(* IEC 61131-3 sources: model-first-plc-agent-ai/results/T2-W-09, 2 files *)

(* ---- a1_code.st ---- *)
FUNCTION_BLOCK TankFillingRuntime
VAR_INPUT
    start : BOOL;
    stop : BOOL;
    LSH : BOOL;
    LSHH : BOOL;
    TimerDuration : TIME;
END_VAR
VAR_OUTPUT
    fill_valve : BOOL;
    discharge_valve : BOOL;
END_VAR
VAR
    x0 : BOOL := TRUE;
    x1 : BOOL := FALSE;
    t1 : BOOL;
    t2 : BOOL;
    timer_done : BOOL := FALSE;
    FillingTimer : TON;
END_VAR

(* Evaluate the start transition from the current situation. *)
t1 := x0 AND start AND NOT stop AND NOT LSHH;

(* Start timing in the same scan that the filling step is entered. *)
FillingTimer(
    IN := x1 OR t1,
    PT := TimerDuration
);

(* The owned condition is neutral on entry to x1. *)
timer_done := x1 AND FillingTimer.Q;

(* Evaluate the return transition before updating the situation. *)
t2 := x1 AND (stop OR LSHH OR timer_done);

IF t1 THEN
    x0 := FALSE;
    x1 := TRUE;
ELSIF t2 THEN
    x0 := TRUE;
    x1 := FALSE;
END_IF;

(* Reset the owned timer immediately when its step is inactive. *)
IF NOT x1 THEN
    FillingTimer(IN := FALSE, PT := TimerDuration);
    timer_done := FALSE;
END_IF;

fill_valve := x1;
discharge_valve := FALSE;

END_FUNCTION_BLOCK

PROGRAM Main
VAR
    StartCommand AT %IX100.0 : BOOL;
    StopCommand AT %IX100.1 : BOOL;
    LSH AT %IX100.2 : BOOL;
    LSHH AT %IX100.3 : BOOL;
    FillValve AT %QX100.0 : BOOL;
    DischargeValve AT %QX100.1 : BOOL;
END_VAR
VAR
    (* Configurable filling duration. *)
    TimerDuration : TIME := T#10s;
    StartEdge : R_TRIG;
    FillingControl : TankFillingRuntime;
END_VAR

StartEdge(CLK := StartCommand);

FillingControl(
    start := StartEdge.Q,
    stop := StopCommand,
    LSH := LSH,
    LSHH := LSHH,
    TimerDuration := TimerDuration
);

FillValve := FillingControl.fill_valve;
DischargeValve := FillingControl.discharge_valve;

END_PROGRAM

(* ---- a2_code.st ---- *)
FUNCTION_BLOCK TankFillingController
VAR_INPUT
    StartCommand : BOOL;
    StopCommand : BOOL;
    LSH : BOOL;
    LSHH : BOOL;
    TimerDuration : TIME;
END_VAR
VAR_OUTPUT
    fill_valve : BOOL;
    discharge_valve : BOOL;
END_VAR
VAR
    StartEdge : R_TRIG;
    FillingTimer : TON;
    start : BOOL;
    stop : BOOL;
    timer_done : BOOL := FALSE;
    x1 : BOOL := FALSE;
END_VAR

StartEdge(CLK := StartCommand);
start := StartEdge.Q;
stop := StopCommand;

IF NOT x1 THEN
    timer_done := FALSE;

    IF start AND NOT stop AND NOT LSHH AND NOT timer_done THEN
        x1 := TRUE;
    END_IF;
END_IF;

FillingTimer(IN := x1, PT := TimerDuration);
timer_done := FillingTimer.Q;

IF stop OR LSHH OR timer_done THEN
    x1 := FALSE;
END_IF;

fill_valve := x1;
discharge_valve := FALSE;

END_FUNCTION_BLOCK

PROGRAM Main
VAR
    StartCommand AT %IX100.0 : BOOL;
    StopCommand AT %IX100.1 : BOOL;
    LSH AT %IX100.2 : BOOL;
    LSHH AT %IX100.3 : BOOL;
    FillValve AT %QX100.0 : BOOL;
    DischargeValve AT %QX100.1 : BOOL;
END_VAR
VAR
    TimerDuration : TIME := T#10s;
    Controller : TankFillingController;
END_VAR

Controller(
    StartCommand := StartCommand,
    StopCommand := StopCommand,
    LSH := LSH,
    LSHH := LSHH,
    TimerDuration := TimerDuration
);

FillValve := Controller.fill_valve;
DischargeValve := Controller.discharge_valve;

END_PROGRAM
